FUNCTION_BLOCK FB_BECKHOFFDRIVE_REF
VAR_INPUT
	stTerminalState			AT %I*:ST_TerminalState;
	stBECKHOFFToPlc		AT %I*:ST_BECKHOFFDRIVETOPLC;
	stPlcToBECKHOFF		AT %Q*:ST_PLCTOBECKHOFFDRIVE;
END_VAR
VAR_OUTPUT

END_VAR
VAR_IN_OUT

END_VAR
VAR

END_VAR

;

END_FUNCTION_BLOCK

(* stored: Version 1.1.0.1, ProductVersion 3.1.4024.15
   POU FB_BECKHOFFDRIVE_REF: Id {73655d98-7033-4df1-889a-0e1f1abc64a6}, SpecialFunc None *)
